Staubli VAL3: do_if.pgx

public program do_if(string x_sKey, num x_nIndex, bool& x_bResult)
  local num l_nType[3]
  local num l_nIndex[3]
  local num l_nValue[3]
  local bool l_bResult1
  local bool l_bDisable1
  local bool l_bResult2
  local bool l_bDisable2
  local bool l_bResult3
  local bool l_bDisable3
  local bool l_bANDOR1
  local bool l_bANDOR2
  local num l_i
begin
  for l_i = 0 to 2
    l_nType[l_i]=progTemp:pProgItem[x_sKey].pProgTemplate[x_nIndex].iIfItem.nSigType[l_i]
    l_nIndex[l_i]=progTemp:pProgItem[x_sKey].pProgTemplate[x_nIndex].iIfItem.nSigIndex[l_i]
    l_nValue[l_i]=progTemp:pProgItem[x_sKey].pProgTemplate[x_nIndex].iIfItem.nValue[l_i]
  endFor

  l_bANDOR1=(progTemp:pProgItem[x_sKey].pProgTemplate[x_nIndex].iIfItem.bANDOR[0]==true)
  l_bANDOR2=(progTemp:pProgItem[x_sKey].pProgTemplate[x_nIndex].iIfItem.bANDOR[1]==true)

  call if_check(l_nType[0],l_nIndex[0],l_nValue[0],l_bResult1,l_bDisable1)
  call if_check(l_nType[1],l_nIndex[1],l_nValue[1],l_bResult2,l_bDisable2)
  call if_check(l_nType[2],l_nIndex[2],l_nValue[2],l_bResult3,l_bDisable3)

  if l_bDisable2
    x_bResult=l_bResult1
  else
    if l_bANDOR1
      x_bResult=(l_bResult1 or l_bResult2)
    else
      x_bResult=(l_bResult1 and l_bResult2)
    endIf

    if l_bDisable3
    else
      if l_bANDOR2
        x_bResult=(x_bResult and (l_bResult2 or l_bResult3))
      else
        x_bResult=x_bResult and (l_bResult2 and l_bResult3)
      endIf
    endIf
  endIf



end
